(* IEC 61131-3 sources: ZPLC/packages/zplc-ide/projects/edge_counter_starter/src, 1 file *)

(* ---- EdgeCounter.st ---- *)
PROGRAM EdgeCounter
VAR_INPUT PulseInput AT %I0.0 : BOOL; Reset AT %I0.1 : BOOL; END_VAR
VAR_OUTPUT CountReached AT %Q0.0 : BOOL; END_VAR
(* Exercise: add a CTU with PV 3: CountReached turns ON on the third rising edge of PulseInput and Reset clears the count. *)
CountReached := FALSE;
END_PROGRAM
